Staubli VAL3: NewApp.pjx

--- NewApp.pjx ---
Parameters version=s8.15.3Cs9_BS3337 stackSize=200000 millimeterUnit=true
Program file=init.pgx
Program file=start.pgx
Program file=stop.pgx
Program file=taskManager.pgx
Program file=stateMachine.pgx
Data file=NewApp.dtx

--- NewApp.dtx ---
public num nState
public num nAlarm
public string sAlarmMsg
public bool bStartCmd
public bool bStopCmd
public bool bPauseCmd
public bool bResetCmd
public bool bRunning
public num nCycleCount
public num nProdCount

--- start.pgx ---
program start()
begin
  //应用入口。SRS 下载后在“应用管理”里设为启动应用即可自动执行。
  call init()

  //核心任务：状态机（优先级高于 HMI）
  taskCreate "stateMachine",50,stateMachine()
  //任务守护：任务异常退出后自动拉起，保证长期运行
  taskCreate "taskManager",20,taskManager()

  //主程序作为心跳，不退出
  do
    delay(1)
  until false
end

--- init.pgx ---
program init()
begin
  //应用初始化：可重复调用（幂等）
  nState=0
  nAlarm=0
  sAlarmMsg=""
  bStartCmd=false
  bStopCmd=false
  bPauseCmd=false
  bResetCmd=false
  bRunning=false
  nCycleCount=0
  nProdCount=0
end

--- stateMachine.pgx ---
program stateMachine()
begin
  //运行状态机
  //  0  初始化
  //  10 空闲（等待启动）
  //  20 运行（执行工艺）
  //  30 暂停
  //  90 故障（报警，等待复位）
  do
    switch nState
      case 0
        //上电/复位后的初始化
        call init()
        nState=10
      break

      case 10
        //空闲：等待启动指令
        bRunning=false
        if bStartCmd
          bStartCmd=false
          nState=20
        endIf
      break

      case 20
        //运行：在这里调用工艺程序
        //  call cycle()
        //  说明：cycle() 是待实现的工艺程序，放在独立的 .pjx 模块里，
        //        通过 Libraries 引用后写作 call <alias>:cycle()
        bRunning=true
        nCycleCount=nCycleCount+1
        //占位：真正的工艺调用接好后删掉这一行
        delay(0.01)
        if bPauseCmd
          bPauseCmd=false
          nState=30
        endIf
        if bStopCmd
          bStopCmd=false
          nState=10
        endIf
      break

      case 30
        //暂停：保持当前位置，等待继续或停止
        bRunning=false
        if bStartCmd
          bStartCmd=false
          nState=20
        endIf
        if bStopCmd
          bStopCmd=false
          nState=10
        endIf
      break

      case 90
        //故障：等待复位
        bRunning=false
        if bResetCmd
          bResetCmd=false
          nAlarm=0
          sAlarmMsg=""
          nState=10
        endIf
      break
    endSwitch
    delay(0)
  until false
end

--- stop.pgx ---
program stop()
begin
  //应用停止时调用：让机器人停在安全状态
  bRunning=false
  nState=0
end

--- taskManager.pgx ---
program taskManager()
begin
  //任务守护：某个任务因通信中断/异常退出后，5 秒后自动拉起
  do
    if taskStatus("stateMachine")!=1
      taskResume("stateMachine",1)
      delay(5)
    endIf
    delay(0)
  until false
end
